Fanuc KAREL source: kd00023.KL

-- PROVISIONAL review KL for V770-1; original PC SHA256 8df127e4788fc0da7e735c68a83ccc2159076b2e34ab84e0588206a559735de5
-- Incomplete behavior may be omitted. Consult companion uncertainty JSON. Do not deploy.
PROGRAM KD00023
%NOLOCKGROUP
VAR
  I : INTEGER
  J : INTEGER
  B : BOOLEAN
  R : REAL
  S : STRING[80]
  SAVED : INTEGER
BEGIN
  -- UNRESOLVED_PC offsets 5-17; opcodes 21,23
  -- UNRESOLVED_PC offsets 22-26; opcodes 7F
END KD00023
